FUNCTION_BLOCK FbFailComposto (* FbFail = alarme de realimentacao OU falha OU intertravamento *)
  (* Standard: 61499-2 *)
  (* Version 1.0, 04/11/2026, Hidryco, Hidryco, 1.0: FbFailOut.value = FbAlarm.value OU Fail OU IlckCond; qualidade do FbAlarm; carimbo de tempo novo quando o valor muda. Usado nos CATs MotorVsBaseNer, MotorBaseNer e ValveBaseNer antes do IThis.FbFail. *)
  PACKAGE SE.Nereda;
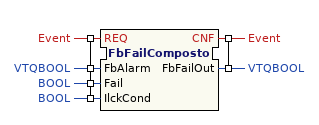
  EVENT_INPUT
    REQ WITH FbAlarm, Fail, IlckCond; (* Recalcula *)
  END_EVENT
  EVENT_OUTPUT
    CNF WITH FbFailOut; (* FbFail composto *)
  END_EVENT
  VAR_INPUT
    FbAlarm : VTQBOOL; (* AlarmStatus do alarme de realimentacao (feedbackFailure) *)
    Fail : BOOL; (* 1 = falha ativa *)
    IlckCond : BOOL; (* 1 = intertravamento ativo *)
  END_VAR
  VAR_OUTPUT
    FbFailOut : VTQBOOL; (* Para o IThis.FbFail *)
  END_VAR
  VAR
    Novo : BOOL; (* Valor calculado *)
  END_VAR
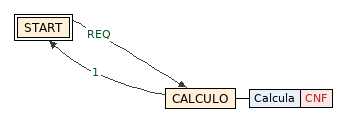
  EC_STATES
    START; (* Estado inicial *)
    CALCULO : Calcula -> CNF; (* Calcula o FbFail *)
  END_STATES
  EC_TRANSITIONS
    START TO CALCULO := REQ;
    CALCULO TO START := 1;
  END_TRANSITIONS
  ALGORITHM Calcula IN ST: (* OU com carimbo de tempo *)
Novo := FbAlarm.value OR Fail OR IlckCond;
IF Novo <> FbFailOut.value THEN
    FbFailOut.timestamp := CURRENT_DT();
END_IF;
FbFailOut.value := Novo;
FbFailOut.quality := FbAlarm.quality;
  END_ALGORITHM
END_FUNCTION_BLOCK
